// ============================================================================
// ST_Station1.scl - 汇川换型改造 工位1 动作机构数据类型定义
// ============================================================================
// 描述:
//   定义 DJ-2026-009 汇川换型改造 工位1 的控制、状态、配置、传感器与执行器结构体.
//   遵循 LSP-905 命名与结构化规范, 支持结构体整块传递 (Struct Chunk Passing).
// ============================================================================

TYPE ST_Station1_Control :
STRUCT
    bAutoEnable     : BOOL;     // 自动运行使能
    bManualStart    : BOOL;     // 手动单步启动
    bReset          : BOOL;     // 故障复位
    bPause          : BOOL;     // 暂停
    bSingleStepMode : BOOL;     // 单步模式
END_STRUCT;
END_TYPE

TYPE ST_Station1_Status :
STRUCT
    iStep           : DINT;     // 当前工步号
    bRunning        : BOOL;     // 运行中
    bDone           : BOOL;     // 本周期动作完成
    bAlarm          : BOOL;     // 站级报警
    iAlarmCode      : DINT;     // 报警代码 (101~199)
    bWaitMaterial   : BOOL;     // 等待来料
    bProcessing     : BOOL;     // 加工中
END_STRUCT;
END_TYPE

TYPE ST_Station1_Config :
STRUCT
    dDebounceMs     : DINT;     // 光电消抖时间 (ms, 默认 100)
    dCylTimeoutMs   : DINT;     // 气缸动作超时时间 (ms, 默认 5000)
    dProcessTimeMs  : DINT;     // 工艺加工延时时间 (ms, 默认 2000)
END_STRUCT;
END_TYPE

TYPE ST_Station1_Sensors :
STRUCT
    bInPosSensor    : BOOL;     // 入料到位光电
    bWorkPosSensor  : BOOL;     // 加工到位光电
END_STRUCT;
END_TYPE

TYPE ST_Station1_Actuators :
STRUCT
    stMotorFwd      : ST_ConveyorMotor; // 进料输送电机
    stCyl1          : ST_Cylinder;      // 夹紧气缸
    stCyl2          : ST_Cylinder;      // 顶升气缸
END_STRUCT;
END_TYPE

TYPE ST_Station1 :
STRUCT
    stControl       : ST_Station1_Control;     // 工位1 控制命令
    stStatus        : ST_Station1_Status;      // 工位1 状态反馈
    stConfig        : ST_Station1_Config;      // 工位1 参数配置
    stSensors       : ST_Station1_Sensors;     // 工位1 传感器输入
    stActuators     : ST_Station1_Actuators;   // 工位1 执行器输出
END_STRUCT;
END_TYPE
